DATA_BLOCK "FRK_PersistAnchors"
{ S7_Optimized_Access := 'TRUE' }
VERSION : 0.1
NON_RETAIN
VAR RETAIN
    RowsA {ExternalAccessible := 'False'; ExternalVisible := 'False'; ExternalWritable := 'False'} : Array[1..17] of "FRK_PersistAnchor";
    RowsB {ExternalAccessible := 'False'; ExternalVisible := 'False'; ExternalWritable := 'False'} : Array[1..17] of "FRK_PersistAnchor";
    SelectedB {ExternalAccessible := 'False'; ExternalVisible := 'False'; ExternalWritable := 'False'} : Array[1..17] of Bool;
    Commissioned {ExternalAccessible := 'False'; ExternalVisible := 'False'; ExternalWritable := 'False'} : Array[1..17] of Bool;
END_VAR
BEGIN
END_DATA_BLOCK
